// TIA Portal V20 export
Screen "Pop-up_StyleConfigRFIDWrite"  641x452
